FUNCTION_BLOCK "Baustein_1"   // FB2222, GRAPH
{ S7_Optimized_Access := 'FALSE' }
VERSION : 0.1
   VAR_INPUT
      INIT_SQ : Bool := false;   // Kette in Initialzustand versetzen
      A_EIN : Bool;
      A_NOT_HALT : Bool;
      Nachfolgendes_Agg_frei : Bool;
      Sensor_vorheriges_Agg : Bool;
      Sensor_Anfang : Bool;   // Öffner
      Sensor_Ende : Bool;   // Öffner
   END_VAR
   VAR_OUTPUT
      Schritt_Nummer : Int;
      Aggregat : Bool;
      Aggregat_frei : Bool;
   END_VAR
   VAR
      HM_FLAM : Array[1..8] of Bool;
      Flanke : Array[1..8] of Bool;
      HM_Agg_Frei : Bool;
      HM_belegt : Bool;
      SWITCH : Array[0..0] of DWord;
      SW_SQTS : Array[0..6] of Byte;
      SW_ADDR : Word := 16#C;
      G7T_0 : GraphTransition;
      G7S_0 : GraphStep;
      PRE_CRIT : Array[0..1] of DWord;
      POST_CRIT : Array[0..0] of DWord;
      TVX : Array[0..2] of Byte;
      TTX : Array[0..2] of Byte;
      TSX : Array[0..2] of Byte;
      S00X : Array[0..2] of Byte;
      SOFFX : Array[0..2] of Byte;
      SONX : Array[0..2] of Byte;
      SAX : Array[0..2] of Byte;
      SERRX : Array[0..7] of Byte;
      SMX : Array[0..7] of Byte;
      S0X : Array[0..7] of Byte;
      S1X : Array[0..7] of Byte;
      S_DISPLAY : Int;   // Interne Anzeige des Ausgangsparameters S_NO
      S_SEL_OLD : Int;   // Vorheriger Wert an S_SEL
      S_DISPIDX : Byte;   // Index des Schritts, der an S_NO anliegt
      T_DISPIDX : Byte;   // Index der Transition, die an T_NO anliegt
      MOPEDGE : Struct
         AUTO : Bool := false;
         MAN : Bool := false;
         TAP : Bool := false;
         TOP : Bool := false;
         ACK_S : Bool := false;
         REG_S : Bool := false;
         T_PREV : Bool := false;
         T_NEXT : Bool := false;
         LOCK : Bool := false;
         SUP : Bool := false;
         ACKREQ : Bool := false;
         SSKIP : Bool := false;
         OFF : Bool := false;
         INIT : Bool := false;
         HALT : Bool := false;
         TMS_HALT : Bool := false;
         OPS_ZERO : Bool := false;
         SACT_DISP : Bool := false;
         SEF_DISP : Bool := false;
         SALL_DISP : Bool := false;
         S_PREV : Bool := false;
         S_NEXT : Bool := false;
         S_SELOK : Bool := false;
         S_ON : Bool := false;
         S_OFF : Bool := false;
         T_PUSH : Bool := false;
         REG : Bool := false;
         ACK : Bool := false;
         IL_PERM : Bool := false;
         T_PERM : Bool := false;
         ILP_MAN : Bool := false;
      END_STRUCT;
      MOP : Struct   // Betriebsart
         AUTO : Bool := true;   // Zustand: Automatischer Betrieb
         MAN : Bool := false;   // Zustand: Handbetrieb
         TAP : Bool := false;   // Zustand: Halbautomatisch/Weiterschalten mit Transition
         TOP : Bool := false;   // Zustand: Halbautomatisch/Ignoriere Transition
         ACK_S : Bool := false;   // Anforderung: Schritt quittieren, der an Parameter S_NO anliegt
         REG_S : Bool := false;   // Anforderung: Schritt registrieren, der an Parameter S_NO anliegt
         T_PREV : Bool := false;   // Anforderung: Vorherige gültige Transition am Parameter T_NO ausgeben
         T_NEXT : Bool := false;   // Anforderung: Nächste gültige Transition am Parameter T_NO ausgeben
         LOCK : Bool := true;   // Zustand: Interlockbearbeitung aktiviert
         SUP : Bool := true;   // Zustand: Supervisionsbearbeitung aktiviert
         ACKREQ : Bool := false;   // Zustand: Quittierung erforderlich
         SSKIP : Bool := false;   // Zustand: "Schritte überspringen" aktiviert
         OFF : Bool := false;   // Anforderung: Alle Schritte deaktivieren
         INIT : Bool := true;   // Anforderung: Kette in Initialzustand schalten
         HALT : Bool := false;   // Zustand: Kette schaltet nicht weiter
         TMS_HALT : Bool := false;   // Zustand: Alle internen Zeiten angehalten
         OPS_ZERO : Bool := false;   // Zustand: Alle mit N, L, D bearbeitete Operanden auf 0 gesetzt
         SACT_DISP : Bool := true;   // Zustand: Nur aktive Schritte anzeigen
         SEF_DISP : Bool := false;   // Zustand: Nur fehlerhafte und gestörte Schritte anzeigen
         SALL_DISP : Bool := false;   // Zustand: Alle Schritte anzeigen
         S_PREV : Bool := false;   // Anforderung: Vorherigen Schritt am Parameter S_NO ausgeben
         S_NEXT : Bool := false;   // Anforderung: Nächsten Schritt am Parameter S_NO ausgeben
         S_SELOK : Bool := false;   // Anforderung: Schrittnummer, die am Parameter S_SEL anliegt, am Parameter S_NO ausgeben
         S_ON : Bool := false;   // Anforderung: Schritt aktivieren, der am Parameter S_NO anliegt
         S_OFF : Bool := false;   // Anforderung: Schritt deaktivieren, der am Parameter S_NO anliegt
         T_PUSH : Bool := false;   // Anforderung: Schaltfreigabe für Transition
         REG : Bool := false;   // Anforderung: Alle Interlock- und Supervisionsfehler registrieren
         ACK : Bool := false;   // Anforderung: Alle Interlock- und Supervisionsfehler quittieren
         IL_PERM : Bool := false;   // Zustand: Permanente Bearbeitung aller Interlocks
         T_PERM : Bool := false;   // Zustand: Permanente Bearbeitung aller Transitionen
         ILP_MAN : Bool := false;   // Zustand: Permanente Bearbeitung aller Interlocks im Handbetrieb
      END_STRUCT;
      TICKS : Struct   // Zeittakte
         DELTA : Time := T#0ms;   // Zeitdifferenz zwischen zwei Zyklen
         OLD : Time := T#0ms;   // 10 ms Taktzählerstand im letzten Zyklus
         NEW : Time := T#0ms;   // 10 ms Taktzählerstand in diesem Zyklus
      END_STRUCT;
      SQ_FLAGS : Struct   // Kettenmerker
         ERR_FLT : Bool := false;   // Sammelfehler Interlock und Supervision
         ERROR : Bool := false;   // Sammelfehler Interlock
         FAULT : Bool := false;   // Sammelfehler Supervision
         RT_FAIL : Bool := false;   // Laufzeitfehler
         NO_SNO : Bool := false;   // Angeforderte Schrittnummer nicht gefunden
         NF_OFL : Bool := false;   // Überlauf: Zu viele Anforderungen ON oder OFF
         SA_OFL : Bool := false;   // Überlauf: Zu viele Schritte aktiv
         TV_OFL : Bool := false;   // Überlauf: Zu viele gültige Transitionen
         MSG_OFL : Bool := false;   // Überlauf: Nicht genügend Systemressourcen fü ALARM_S
         NO_SWI : Bool := false;   // Nicht Schalten in diesem Zyklus
         CYC_OP : Bool := false;   // Zyklische Bearbeitung der Kette nach Initialisierung
         AS_MSG : Bool := true;   // Meldungen zur Laufzeit durch Anweisung aktiviert oder deaktiviert
         AS_SEND : Bool := false;   // Meldungen von WR_USMSG senden oder nur in Diagnosepuffer eintragen
         SQ_BUSY : Bool := false;   // Interner Flankenmerker für Vorgangsbearbeitung
         SA_BUSY : Bool := false;   // Interner Flankenmerker für Vorgangsbearbeitung
         AS_SIG : Bool := false;   // Flankenmerker für Meldungen von Alarm_S und Alarm_SQ
      END_STRUCT;
      S_PTR : DWord := 16#450;
      S_PTR2 : DWord := 16#0;
      S_PTR3 : DWord := 16#D50;
      S_PTR4 : DWord := 16#D10;
      T_PTR : DWord := 16#CD0;
      C_AR2 : DWord := 16#0;
      M_FBDB : DWord := 16#8AE0000;
      M_SNO : Word := 16#4;
      M_EVID : Word := 16#0;
      M_EVIL : C_Alarm_s;
      M_EVSV : C_Alarm_s;
      M_EV : DWord := 16#C30;
      CRIT : Array[0..31] of Bool;
      S_START : Byte := 16#0;
      S_IDX : Byte := 16#0;
      S_INT : Int := 72;
      S_TMP : Byte := 16#0;
      T_START : Byte := 16#0;
      T_IDX : Byte := 16#0;
      T_TMP : Byte := 16#0;
      T_TMP2 : Byte := 16#00;
      TV_POT : Byte := 16#02;
      RETURN1 : Byte := 16#0;
      RETURN2 : Byte := 16#0;
      SINI : Array[0..2] of Byte;
      LSTT : Array[0..6] of Byte;
      ATAJ : Array[0..6] of Byte;
      ATAB : Array[0..6] of Byte;
      PSTT : Array[0..6] of Byte;
      NSTT : Array[0..6] of Byte;
      ASSJ : Array[0..6] of Byte;
      ASSB : Array[0..6] of Byte;
      PTTS : Array[0..6] of Byte;
      NTTS : Array[0..6] of Byte;
      PRE_CNT : Word := 16#2;
      POST_CNT : Word := 16#1;
      ADR_COND : Word := 16#0;
      MAX_TVAL : Byte := 16#1;
      MAX_SACT : Byte := 16#1;
      MAX_CRIT : Byte := 16#4;
      T_CNT : Byte := 16#6;
      SUP_CNT : Byte := 16#0;
      LOCK_CNT : Byte := 16#5;
      S_CNT : Byte := 16#6;
      SQ_CNT : Byte := 16#1;
      PRS_INPAR : DWord := 16#40000000;
      PRS_OUTPAR : DWord := 16#0;
      GC_FLAGS : Struct
         T_MACH : Byte := 16#EB;
         COND_ED : Byte := 16#E2;
         W_LEVEL : Byte := 16#D5;
         FB_IF : Byte := 16#FA;
         AS_MSG : Word := 16#404;
         SSB : Word := 16#108;
         DILG : Word := 16#27E;
         ADDR_T0 : Word := 16#1A;
         CRIT_AVAIL : Bool := false;
         SSKIP_AVAIL : Bool := true;
         SSKIP_ON : Bool := false;
         ACK_REQ : Bool := false;
         SYNC_AVAIL : Bool := true;
         ILP_MAN : Bool := false;
         SWM_LOCKED : Bool := false;
         SAVE_SW : Bool := true;
      END_STRUCT;
      G7_FBMARK : Byte := 16#3C;
      G7_RELEASE : Byte := 16#3C;
      G7_ID2 : Byte := 16#37;
      G7_ID1 : Byte := 16#47;
   END_VAR
   // SW_SQTS[0] := 16#1;
   // TVX[0] := 16#1;
   // TTX[0] := 16#1;
   // TSX[0] := 16#1;
   // S00X[0] := 16#1;
   // SOFFX[0] := 16#1;
   // SONX[0] := 16#1;
   // SAX[0] := 16#1;
   // SERRX[0] := 16#1;
   // SMX[0] := 16#1;
   // S0X[0] := 16#1;
   // S1X[0] := 16#1;
   // SINI[0] := 16#2;
   // SINI[1] := 16#1;
   // SINI[2] := 0;
   // LSTT[0] := 0;
   // LSTT[1] := 0;
   // LSTT[2] := 0;
   // LSTT[3] := 0;
   // LSTT[4] := 0;
   // LSTT[5] := 0;
   // LSTT[6] := 16#1;
   // ATAJ[0] := 0;
   // ATAJ[1] := 16#1;
   // ATAJ[2] := 16#2;
   // ATAJ[3] := 16#3;
   // ATAJ[4] := 16#4;
   // ATAJ[5] := 16#5;
   // ATAJ[6] := 16#6;
   // ATAB[0] := 0;
   // ATAB[1] := 16#1;
   // ATAB[2] := 16#2;
   // ATAB[3] := 16#3;
   // ATAB[4] := 16#4;
   // ATAB[5] := 16#5;
   // ATAB[6] := 16#6;
   // PSTT[0] := 0;
   // PSTT[1] := 16#1;
   // PSTT[2] := 16#2;
   // PSTT[3] := 16#3;
   // PSTT[4] := 16#4;
   // PSTT[5] := 16#5;
   // PSTT[6] := 16#6;
   // NSTT[0] := 16#1;
   // NSTT[1] := 16#2;
   // NSTT[2] := 16#3;
   // NSTT[3] := 16#4;
   // NSTT[4] := 16#5;
   // NSTT[5] := 16#6;
   // NSTT[6] := 16#1;
   // ASSJ[0] := 0;
   // ASSJ[1] := 16#1;
   // ASSJ[2] := 16#2;
   // ASSJ[3] := 16#3;
   // ASSJ[4] := 16#4;
   // ASSJ[5] := 16#5;
   // ASSJ[6] := 16#6;
   // ASSB[0] := 0;
   // ASSB[1] := 16#1;
   // ASSB[2] := 16#2;
   // ASSB[3] := 16#3;
   // ASSB[4] := 16#4;
   // ASSB[5] := 16#5;
   // ASSB[6] := 16#6;
   // PTTS[0] := 0;
   // PTTS[2] := 16#1;
   // PTTS[3] := 16#2;
   // PTTS[4] := 16#3;
   // PTTS[5] := 16#4;
   // PTTS[6] := 16#5;
   // NTTS[0] := 0;
   // NTTS[1] := 16#1;
   // NTTS[2] := 16#2;
   // NTTS[3] := 16#3;
   // NTTS[4] := 16#4;
   // NTTS[5] := 16#5;
   // NTTS[6] := 16#6;
BEGIN
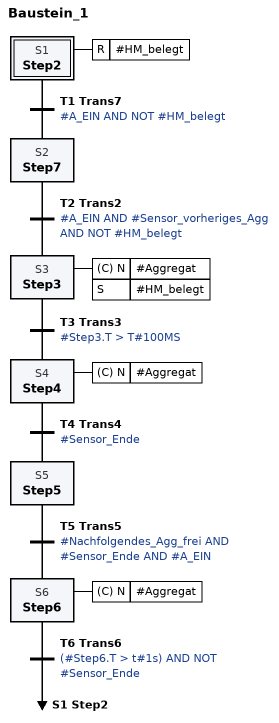
   // permanent pre-instructions
   NETWORK 1
      #HM_Agg_Frei := NOT #HM_belegt;
      #Aggregat_frei := NOT #HM_belegt;
   NETWORK 2
   TITLE = Ausgabe Schrittnummer
      #Schritt_Nummer := #S_DISPLAY;

   // sequencer 1
   INITIAL_STEP Step2:   // S1
      interlock C := NOT #A_NOT_HALT;
      // Warten auf Start
              R    #HM_belegt
   END_STEP
   TRANSITION Trans7 FROM Step2 TO Step7   // T1
      := #A_EIN AND NOT #HM_belegt;
   END_TRANSITION
   STEP Step4:   // S4
      interlock C := NOT #A_NOT_HALT;
      // Einfahrt bis Ende
      (C)     N    #Aggregat
   END_STEP
   TRANSITION Trans4 FROM Step4 TO Step5   // T4
      := #Sensor_Ende;
   END_TRANSITION
   STEP Step5:   // S5
      interlock C := NOT #A_NOT_HALT;
      // Warten auf Ausfahrt
   END_STEP
   TRANSITION Trans5 FROM Step5 TO Step6   // T5
      := #Nachfolgendes_Agg_frei AND #Sensor_Ende AND #A_EIN;
   END_TRANSITION
   STEP Step6:   // S6
      interlock C := NOT #A_NOT_HALT;
      // Ausfahrt bis Ende
      (C)     N    #Aggregat
   END_STEP
   TRANSITION Trans6 FROM Step6 TO Step2   // T6, jump
      := (#Step6.T > t#1s) AND NOT #Sensor_Ende;
   END_TRANSITION
   STEP Step3:   // S3
      interlock C := NOT #A_NOT_HALT;
      // Einfahrt Start
      (C)     N    #Aggregat
              S    #HM_belegt
   END_STEP
   TRANSITION Trans3 FROM Step3 TO Step4   // T3
      := #Step3.T > T#100MS;
   END_TRANSITION
   STEP Step7:   // S2
   END_STEP
   TRANSITION Trans2 FROM Step7 TO Step3   // T2
      := #A_EIN AND #Sensor_vorheriges_Agg AND NOT #HM_belegt;
   END_TRANSITION
END_FUNCTION_BLOCK